// TIA Portal V21 export
VBScript "CheckPump"  Type=Sub
  If SmartTags("PumpSpeed") > 100 Then
    ShowSystemAlarm "Pump speed high"
  End If
